Fanuc KAREL source: kt00474.KL

-- PROVISIONAL review KL for V770-1; original PC SHA256 9d7a969db0a5c335791845e3075033f31ac5b3a96d8877cfd7421063d244559d
-- Incomplete behavior may be omitted. Consult companion uncertainty JSON. Do not deploy.
PROGRAM KT00474
%NOLOCKGROUP
-- UNRESOLVED_DECL P1 type=000101
-- UNRESOLVED_DECL P2 type=000101
-- UNRESOLVED_DECL OUT type=000101
BEGIN
  -- UNRESOLVED_PC offsets 5-29; opcodes 49,49,60,4A
  -- UNRESOLVED_PC offsets 34-38; opcodes 7F
END KT00474
